(* IEC 61131-3 sources: IEC61131-3_ST_SCL_Mutation_Generator/Tests/mutatedCode_fibonacci_number_m, 23 files *)

(* ---- M1349.st ---- *)
FUNCTION_BLOCK "FB_Fibonacci_Calculator"
{ S7_Optimized_Access := 'FALSE' }
VERSION : 1.0

VAR_INPUT
    N : DInt := 5;
END_VAR

VAR_OUTPUT
    O : DInt := 1;
END_VAR

VAR
    F1 : DInt := 1;    // Fib(k-2) at the end of the calculation
    F2 : DInt := 1;    // Fib(k-1) at the end of the calculation
    CNT : DInt := 2;   // Index of the last computed term
END_VAR

BEGIN

    // Start values: Fib(1) = Fib(2) = 1
    #F1 := 1;
    #F2 := 1;
    #O := 1;

    IF #N >= 2 THEN (* MUTATED: REL_OP_REPLACE *)
        // Edge case: N <= 2 returns 1
        #CNT := #N;
    ELSE
        #CNT := 2;
        WHILE #CNT < #N DO
            #CNT := #CNT + 1;

            // Saturation arithmetic: result would exceed INT range
            IF (#F1 + #F2) > 32767 THEN
                #O := 32767;
                EXIT;
            END_IF;

            #O := #F1 + #F2;

            // Shift the window only if another term is still needed,
            // so that at the end O = F1 + F2
            IF #CNT < #N THEN
                #F1 := #F2;
                #F2 := #O;
            END_IF;
        END_WHILE;
    END_IF;

    // Final saturation guard
    IF (#O > 32767) OR (#O < 0) THEN
        #O := 32767;
    END_IF;

    //#ASSERT O >= 0 AND O <= 32767
    //#ASSERT F1 <= 32767 AND F2 <= 32767
    //#ASSERT CNT <= N

END_FUNCTION_BLOCK

(* ---- M1350.st ---- *)
FUNCTION_BLOCK "FB_Fibonacci_Calculator"
{ S7_Optimized_Access := 'FALSE' }
VERSION : 1.0

VAR_INPUT
    N : DInt := 5;
END_VAR

VAR_OUTPUT
    O : DInt := 1;
END_VAR

VAR
    F1 : DInt := 1;    // Fib(k-2) at the end of the calculation
    F2 : DInt := 1;    // Fib(k-1) at the end of the calculation
    CNT : DInt := 2;   // Index of the last computed term
END_VAR

BEGIN

    // Start values: Fib(1) = Fib(2) = 1
    #F1 := 1;
    #F2 := 1;
    #O := 1;

    IF #N <= 2 THEN
        // Edge case: N <= 2 returns 1
        #CNT := #N;
    ELSE
        #CNT := 2;
        WHILE #CNT > #N DO (* MUTATED: REL_OP_REPLACE *)
            #CNT := #CNT + 1;

            // Saturation arithmetic: result would exceed INT range
            IF (#F1 + #F2) > 32767 THEN
                #O := 32767;
                EXIT;
            END_IF;

            #O := #F1 + #F2;

            // Shift the window only if another term is still needed,
            // so that at the end O = F1 + F2
            IF #CNT < #N THEN
                #F1 := #F2;
                #F2 := #O;
            END_IF;
        END_WHILE;
    END_IF;

    // Final saturation guard
    IF (#O > 32767) OR (#O < 0) THEN
        #O := 32767;
    END_IF;

    //#ASSERT O >= 0 AND O <= 32767
    //#ASSERT F1 <= 32767 AND F2 <= 32767
    //#ASSERT CNT <= N

END_FUNCTION_BLOCK

(* ---- M1351.st ---- *)
FUNCTION_BLOCK "FB_Fibonacci_Calculator"
{ S7_Optimized_Access := 'FALSE' }
VERSION : 1.0

VAR_INPUT
    N : DInt := 5;
END_VAR

VAR_OUTPUT
    O : DInt := 1;
END_VAR

VAR
    F1 : DInt := 1;    // Fib(k-2) at the end of the calculation
    F2 : DInt := 1;    // Fib(k-1) at the end of the calculation
    CNT : DInt := 2;   // Index of the last computed term
END_VAR

BEGIN

    // Start values: Fib(1) = Fib(2) = 1
    #F1 := 1;
    #F2 := 1;
    #O := 1;

    IF #N <= 2 THEN
        // Edge case: N <= 2 returns 1
        #CNT := #N;
    ELSE
        #CNT := 2;
        WHILE #CNT < #N DO
            #CNT := #CNT + 1;

            // Saturation arithmetic: result would exceed INT range
            IF (#F1 + #F2) < 32767 THEN (* MUTATED: REL_OP_REPLACE *)
                #O := 32767;
                EXIT;
            END_IF;

            #O := #F1 + #F2;

            // Shift the window only if another term is still needed,
            // so that at the end O = F1 + F2
            IF #CNT < #N THEN
                #F1 := #F2;
                #F2 := #O;
            END_IF;
        END_WHILE;
    END_IF;

    // Final saturation guard
    IF (#O > 32767) OR (#O < 0) THEN
        #O := 32767;
    END_IF;

    //#ASSERT O >= 0 AND O <= 32767
    //#ASSERT F1 <= 32767 AND F2 <= 32767
    //#ASSERT CNT <= N

END_FUNCTION_BLOCK

(* ---- M1352.st ---- *)
FUNCTION_BLOCK "FB_Fibonacci_Calculator"
{ S7_Optimized_Access := 'FALSE' }
VERSION : 1.0

VAR_INPUT
    N : DInt := 5;
END_VAR

VAR_OUTPUT
    O : DInt := 1;
END_VAR

VAR
    F1 : DInt := 1;    // Fib(k-2) at the end of the calculation
    F2 : DInt := 1;    // Fib(k-1) at the end of the calculation
    CNT : DInt := 2;   // Index of the last computed term
END_VAR

BEGIN

    // Start values: Fib(1) = Fib(2) = 1
    #F1 := 1;
    #F2 := 1;
    #O := 1;

    IF #N <= 2 THEN
        // Edge case: N <= 2 returns 1
        #CNT := #N;
    ELSE
        #CNT := 2;
        WHILE #CNT < #N DO
            #CNT := #CNT + 1;

            // Saturation arithmetic: result would exceed INT range
            IF (#F1 + #F2) > 32767 THEN
                #O := 32767;
                EXIT;
            END_IF;

            #O := #F1 + #F2;

            // Shift the window only if another term is still needed,
            // so that at the end O = F1 + F2
            IF #CNT > #N THEN (* MUTATED: REL_OP_REPLACE *)
                #F1 := #F2;
                #F2 := #O;
            END_IF;
        END_WHILE;
    END_IF;

    // Final saturation guard
    IF (#O > 32767) OR (#O < 0) THEN
        #O := 32767;
    END_IF;

    //#ASSERT O >= 0 AND O <= 32767
    //#ASSERT F1 <= 32767 AND F2 <= 32767
    //#ASSERT CNT <= N

END_FUNCTION_BLOCK

(* ---- M1353.st ---- *)
FUNCTION_BLOCK "FB_Fibonacci_Calculator"
{ S7_Optimized_Access := 'FALSE' }
VERSION : 1.0

VAR_INPUT
    N : DInt := 5;
END_VAR

VAR_OUTPUT
    O : DInt := 1;
END_VAR

VAR
    F1 : DInt := 1;    // Fib(k-2) at the end of the calculation
    F2 : DInt := 1;    // Fib(k-1) at the end of the calculation
    CNT : DInt := 2;   // Index of the last computed term
END_VAR

BEGIN

    // Start values: Fib(1) = Fib(2) = 1
    #F1 := 1;
    #F2 := 1;
    #O := 1;

    IF #N <= 2 THEN
        // Edge case: N <= 2 returns 1
        #CNT := #N;
    ELSE
        #CNT := 2;
        WHILE #CNT < #N DO
            #CNT := #CNT + 1;

            // Saturation arithmetic: result would exceed INT range
            IF (#F1 + #F2) > 32767 THEN
                #O := 32767;
                EXIT;
            END_IF;

            #O := #F1 + #F2;

            // Shift the window only if another term is still needed,
            // so that at the end O = F1 + F2
            IF #CNT < #N THEN
                #F1 := #F2;
                #F2 := #O;
            END_IF;
        END_WHILE;
    END_IF;

    // Final saturation guard
    IF (#O < 32767) OR (#O < 0) THEN (* MUTATED: REL_OP_REPLACE *)
        #O := 32767;
    END_IF;

    //#ASSERT O >= 0 AND O <= 32767
    //#ASSERT F1 <= 32767 AND F2 <= 32767
    //#ASSERT CNT <= N

END_FUNCTION_BLOCK

(* ---- M1354.st ---- *)
FUNCTION_BLOCK "FB_Fibonacci_Calculator"
{ S7_Optimized_Access := 'FALSE' }
VERSION : 1.0

VAR_INPUT
    N : DInt := 5;
END_VAR

VAR_OUTPUT
    O : DInt := 1;
END_VAR

VAR
    F1 : DInt := 1;    // Fib(k-2) at the end of the calculation
    F2 : DInt := 1;    // Fib(k-1) at the end of the calculation
    CNT : DInt := 2;   // Index of the last computed term
END_VAR

BEGIN

    // Start values: Fib(1) = Fib(2) = 1
    #F1 := 1;
    #F2 := 1;
    #O := 1;

    IF #N <= 2 THEN
        // Edge case: N <= 2 returns 1
        #CNT := #N;
    ELSE
        #CNT := 2;
        WHILE #CNT < #N DO
            #CNT := #CNT + 1;

            // Saturation arithmetic: result would exceed INT range
            IF (#F1 + #F2) > 32767 THEN
                #O := 32767;
                EXIT;
            END_IF;

            #O := #F1 + #F2;

            // Shift the window only if another term is still needed,
            // so that at the end O = F1 + F2
            IF #CNT < #N THEN
                #F1 := #F2;
                #F2 := #O;
            END_IF;
        END_WHILE;
    END_IF;

    // Final saturation guard
    IF (#O > 32767) OR (#O > 0) THEN (* MUTATED: REL_OP_REPLACE *)
        #O := 32767;
    END_IF;

    //#ASSERT O >= 0 AND O <= 32767
    //#ASSERT F1 <= 32767 AND F2 <= 32767
    //#ASSERT CNT <= N

END_FUNCTION_BLOCK

(* ---- M1355.st ---- *)
FUNCTION_BLOCK "FB_Fibonacci_Calculator"
{ S7_Optimized_Access := 'FALSE' }
VERSION : 1.0

VAR_INPUT
    N : DInt := 5;
END_VAR

VAR_OUTPUT
    O : DInt := 1;
END_VAR

VAR
    F1 : DInt := 1;    // Fib(k-2) at the end of the calculation
    F2 : DInt := 1;    // Fib(k-1) at the end of the calculation
    CNT : DInt := 2;   // Index of the last computed term
END_VAR

BEGIN

    // Start values: Fib(1) = Fib(2) = 1
    #F1 := 1;
    #F2 := 1;
    #O := 1;

    IF #N <= 2 THEN
        // Edge case: N <= 2 returns 1
        #CNT := #N;
    ELSE
        #CNT := 2;
        WHILE #CNT < #N DO
            #CNT := #CNT + 1;

            // Saturation arithmetic: result would exceed INT range
            IF (#F1 + #F2) > 32767 THEN
                #O := 32767;
                EXIT;
            END_IF;

            #O := #F1 + #F2;

            // Shift the window only if another term is still needed,
            // so that at the end O = F1 + F2
            IF #CNT < #N THEN
                #F1 := #F2;
                #F2 := #O;
            END_IF;
        END_WHILE;
    END_IF;

    // Final saturation guard
    IF (#O > 32767) AND (#O < 0) THEN (* MUTATED: LOGICAL_OP_REPLACE *)
        #O := 32767;
    END_IF;

    //#ASSERT O >= 0 AND O <= 32767
    //#ASSERT F1 <= 32767 AND F2 <= 32767
    //#ASSERT CNT <= N

END_FUNCTION_BLOCK

(* ---- M1356.st ---- *)
FUNCTION_BLOCK "FB_Fibonacci_Calculator"
{ S7_Optimized_Access := 'FALSE' }
VERSION : 1.0

VAR_INPUT
    N : DInt := 5;
END_VAR

VAR_OUTPUT
    O : DInt := 1;
END_VAR

VAR
    F1 : DInt := 1;    // Fib(k-2) at the end of the calculation
    F2 : DInt := 1;    // Fib(k-1) at the end of the calculation
    CNT : DInt := 2;   // Index of the last computed term
END_VAR

BEGIN

    // Start values: Fib(1) = Fib(2) = 1
    #F1 := 1;
    #F2 := 1;
    #O := 1;

    IF #N <= 2 THEN
        // Edge case: N <= 2 returns 1
        #CNT := #N;
    ELSE
        #CNT := 2;
        WHILE #CNT < #N DO
            #CNT := #CNT - 1; (* MUTATED: ARITH_OP_REPLACE *)

            // Saturation arithmetic: result would exceed INT range
            IF (#F1 + #F2) > 32767 THEN
                #O := 32767;
                EXIT;
            END_IF;

            #O := #F1 + #F2;

            // Shift the window only if another term is still needed,
            // so that at the end O = F1 + F2
            IF #CNT < #N THEN
                #F1 := #F2;
                #F2 := #O;
            END_IF;
        END_WHILE;
    END_IF;

    // Final saturation guard
    IF (#O > 32767) OR (#O < 0) THEN
        #O := 32767;
    END_IF;

    //#ASSERT O >= 0 AND O <= 32767
    //#ASSERT F1 <= 32767 AND F2 <= 32767
    //#ASSERT CNT <= N

END_FUNCTION_BLOCK

(* ---- M1357.st ---- *)
FUNCTION_BLOCK "FB_Fibonacci_Calculator"
{ S7_Optimized_Access := 'FALSE' }
VERSION : 1.0

VAR_INPUT
    N : DInt := 5;
END_VAR

VAR_OUTPUT
    O : DInt := 1;
END_VAR

VAR
    F1 : DInt := 1;    // Fib(k-2) at the end of the calculation
    F2 : DInt := 1;    // Fib(k-1) at the end of the calculation
    CNT : DInt := 2;   // Index of the last computed term
END_VAR

BEGIN

    // Start values: Fib(1) = Fib(2) = 1
    #F1 := 2; (* MUTATED: CONST_VALUE_REPLACE *)
    #F2 := 1;
    #O := 1;

    IF #N <= 2 THEN
        // Edge case: N <= 2 returns 1
        #CNT := #N;
    ELSE
        #CNT := 2;
        WHILE #CNT < #N DO
            #CNT := #CNT + 1;

            // Saturation arithmetic: result would exceed INT range
            IF (#F1 + #F2) > 32767 THEN
                #O := 32767;
                EXIT;
            END_IF;

            #O := #F1 + #F2;

            // Shift the window only if another term is still needed,
            // so that at the end O = F1 + F2
            IF #CNT < #N THEN
                #F1 := #F2;
                #F2 := #O;
            END_IF;
        END_WHILE;
    END_IF;

    // Final saturation guard
    IF (#O > 32767) OR (#O < 0) THEN
        #O := 32767;
    END_IF;

    //#ASSERT O >= 0 AND O <= 32767
    //#ASSERT F1 <= 32767 AND F2 <= 32767
    //#ASSERT CNT <= N

END_FUNCTION_BLOCK

(* ---- M1358.st ---- *)
FUNCTION_BLOCK "FB_Fibonacci_Calculator"
{ S7_Optimized_Access := 'FALSE' }
VERSION : 1.0

VAR_INPUT
    N : DInt := 5;
END_VAR

VAR_OUTPUT
    O : DInt := 1;
END_VAR

VAR
    F1 : DInt := 1;    // Fib(k-2) at the end of the calculation
    F2 : DInt := 1;    // Fib(k-1) at the end of the calculation
    CNT : DInt := 2;   // Index of the last computed term
END_VAR

BEGIN

    // Start values: Fib(1) = Fib(2) = 1
    #F1 := 1;
    #F2 := 2; (* MUTATED: CONST_VALUE_REPLACE *)
    #O := 1;

    IF #N <= 2 THEN
        // Edge case: N <= 2 returns 1
        #CNT := #N;
    ELSE
        #CNT := 2;
        WHILE #CNT < #N DO
            #CNT := #CNT + 1;

            // Saturation arithmetic: result would exceed INT range
            IF (#F1 + #F2) > 32767 THEN
                #O := 32767;
                EXIT;
            END_IF;

            #O := #F1 + #F2;

            // Shift the window only if another term is still needed,
            // so that at the end O = F1 + F2
            IF #CNT < #N THEN
                #F1 := #F2;
                #F2 := #O;
            END_IF;
        END_WHILE;
    END_IF;

    // Final saturation guard
    IF (#O > 32767) OR (#O < 0) THEN
        #O := 32767;
    END_IF;

    //#ASSERT O >= 0 AND O <= 32767
    //#ASSERT F1 <= 32767 AND F2 <= 32767
    //#ASSERT CNT <= N

END_FUNCTION_BLOCK

(* ---- M1359.st ---- *)
FUNCTION_BLOCK "FB_Fibonacci_Calculator"
{ S7_Optimized_Access := 'FALSE' }
VERSION : 1.0

VAR_INPUT
    N : DInt := 5;
END_VAR

VAR_OUTPUT
    O : DInt := 1;
END_VAR

VAR
    F1 : DInt := 1;    // Fib(k-2) at the end of the calculation
    F2 : DInt := 1;    // Fib(k-1) at the end of the calculation
    CNT : DInt := 2;   // Index of the last computed term
END_VAR

BEGIN

    // Start values: Fib(1) = Fib(2) = 1
    #F1 := 1;
    #F2 := 1;
    #O := 2; (* MUTATED: CONST_VALUE_REPLACE *)

    IF #N <= 2 THEN
        // Edge case: N <= 2 returns 1
        #CNT := #N;
    ELSE
        #CNT := 2;
        WHILE #CNT < #N DO
            #CNT := #CNT + 1;

            // Saturation arithmetic: result would exceed INT range
            IF (#F1 + #F2) > 32767 THEN
                #O := 32767;
                EXIT;
            END_IF;

            #O := #F1 + #F2;

            // Shift the window only if another term is still needed,
            // so that at the end O = F1 + F2
            IF #CNT < #N THEN
                #F1 := #F2;
                #F2 := #O;
            END_IF;
        END_WHILE;
    END_IF;

    // Final saturation guard
    IF (#O > 32767) OR (#O < 0) THEN
        #O := 32767;
    END_IF;

    //#ASSERT O >= 0 AND O <= 32767
    //#ASSERT F1 <= 32767 AND F2 <= 32767
    //#ASSERT CNT <= N

END_FUNCTION_BLOCK

(* ---- M1360.st ---- *)
FUNCTION_BLOCK "FB_Fibonacci_Calculator"
{ S7_Optimized_Access := 'FALSE' }
VERSION : 1.0

VAR_INPUT
    N : DInt := 5;
END_VAR

VAR_OUTPUT
    O : DInt := 1;
END_VAR

VAR
    F1 : DInt := 1;    // Fib(k-2) at the end of the calculation
    F2 : DInt := 1;    // Fib(k-1) at the end of the calculation
    CNT : DInt := 2;   // Index of the last computed term
END_VAR

BEGIN

    // Start values: Fib(1) = Fib(2) = 1
    #F1 := 1;
    #F2 := 1;
    #O := 1;

    IF #N <= 3 THEN (* MUTATED: CONST_VALUE_REPLACE *)
        // Edge case: N <= 2 returns 1
        #CNT := #N;
    ELSE
        #CNT := 2;
        WHILE #CNT < #N DO
            #CNT := #CNT + 1;

            // Saturation arithmetic: result would exceed INT range
            IF (#F1 + #F2) > 32767 THEN
                #O := 32767;
                EXIT;
            END_IF;

            #O := #F1 + #F2;

            // Shift the window only if another term is still needed,
            // so that at the end O = F1 + F2
            IF #CNT < #N THEN
                #F1 := #F2;
                #F2 := #O;
            END_IF;
        END_WHILE;
    END_IF;

    // Final saturation guard
    IF (#O > 32767) OR (#O < 0) THEN
        #O := 32767;
    END_IF;

    //#ASSERT O >= 0 AND O <= 32767
    //#ASSERT F1 <= 32767 AND F2 <= 32767
    //#ASSERT CNT <= N

END_FUNCTION_BLOCK

(* ---- M1361.st ---- *)
FUNCTION_BLOCK "FB_Fibonacci_Calculator"
{ S7_Optimized_Access := 'FALSE' }
VERSION : 1.0

VAR_INPUT
    N : DInt := 5;
END_VAR

VAR_OUTPUT
    O : DInt := 1;
END_VAR

VAR
    F1 : DInt := 1;    // Fib(k-2) at the end of the calculation
    F2 : DInt := 1;    // Fib(k-1) at the end of the calculation
    CNT : DInt := 2;   // Index of the last computed term
END_VAR

BEGIN

    // Start values: Fib(1) = Fib(2) = 1
    #F1 := 1;
    #F2 := 1;
    #O := 1;

    IF #N <= 2 THEN
        // Edge case: N <= 2 returns 1
        #CNT := #N;
    ELSE
        #CNT := 3; (* MUTATED: CONST_VALUE_REPLACE *)
        WHILE #CNT < #N DO
            #CNT := #CNT + 1;

            // Saturation arithmetic: result would exceed INT range
            IF (#F1 + #F2) > 32767 THEN
                #O := 32767;
                EXIT;
            END_IF;

            #O := #F1 + #F2;

            // Shift the window only if another term is still needed,
            // so that at the end O = F1 + F2
            IF #CNT < #N THEN
                #F1 := #F2;
                #F2 := #O;
            END_IF;
        END_WHILE;
    END_IF;

    // Final saturation guard
    IF (#O > 32767) OR (#O < 0) THEN
        #O := 32767;
    END_IF;

    //#ASSERT O >= 0 AND O <= 32767
    //#ASSERT F1 <= 32767 AND F2 <= 32767
    //#ASSERT CNT <= N

END_FUNCTION_BLOCK

(* ---- M1362.st ---- *)
FUNCTION_BLOCK "FB_Fibonacci_Calculator"
{ S7_Optimized_Access := 'FALSE' }
VERSION : 1.0

VAR_INPUT
    N : DInt := 5;
END_VAR

VAR_OUTPUT
    O : DInt := 1;
END_VAR

VAR
    F1 : DInt := 1;    // Fib(k-2) at the end of the calculation
    F2 : DInt := 1;    // Fib(k-1) at the end of the calculation
    CNT : DInt := 2;   // Index of the last computed term
END_VAR

BEGIN

    // Start values: Fib(1) = Fib(2) = 1
    #F1 := 1;
    #F2 := 1;
    #O := 1;

    IF #N <= 2 THEN
        // Edge case: N <= 2 returns 1
        #CNT := #N;
    ELSE
        #CNT := 2;
        WHILE #CNT < #N DO
            #CNT := #CNT + 2; (* MUTATED: CONST_VALUE_REPLACE *)

            // Saturation arithmetic: result would exceed INT range
            IF (#F1 + #F2) > 32767 THEN
                #O := 32767;
                EXIT;
            END_IF;

            #O := #F1 + #F2;

            // Shift the window only if another term is still needed,
            // so that at the end O = F1 + F2
            IF #CNT < #N THEN
                #F1 := #F2;
                #F2 := #O;
            END_IF;
        END_WHILE;
    END_IF;

    // Final saturation guard
    IF (#O > 32767) OR (#O < 0) THEN
        #O := 32767;
    END_IF;

    //#ASSERT O >= 0 AND O <= 32767
    //#ASSERT F1 <= 32767 AND F2 <= 32767
    //#ASSERT CNT <= N

END_FUNCTION_BLOCK

(* ---- M1363.st ---- *)
FUNCTION_BLOCK "FB_Fibonacci_Calculator"
{ S7_Optimized_Access := 'FALSE' }
VERSION : 1.0

VAR_INPUT
    N : DInt := 5;
END_VAR

VAR_OUTPUT
    O : DInt := 1;
END_VAR

VAR
    F1 : DInt := 1;    // Fib(k-2) at the end of the calculation
    F2 : DInt := 1;    // Fib(k-1) at the end of the calculation
    CNT : DInt := 2;   // Index of the last computed term
END_VAR

BEGIN

    // Start values: Fib(1) = Fib(2) = 1
    #F1 := 1;
    #F2 := 1;
    #O := 1;

    IF #N <= 2 THEN
        // Edge case: N <= 2 returns 1
        #CNT := #N;
    ELSE
        #CNT := 2;
        WHILE #CNT < #N DO
            #CNT := #CNT + 1;

            // Saturation arithmetic: result would exceed INT range
            IF (#F1 + #F2) > 32768 THEN (* MUTATED: CONST_VALUE_REPLACE *)
                #O := 32767;
                EXIT;
            END_IF;

            #O := #F1 + #F2;

            // Shift the window only if another term is still needed,
            // so that at the end O = F1 + F2
            IF #CNT < #N THEN
                #F1 := #F2;
                #F2 := #O;
            END_IF;
        END_WHILE;
    END_IF;

    // Final saturation guard
    IF (#O > 32767) OR (#O < 0) THEN
        #O := 32767;
    END_IF;

    //#ASSERT O >= 0 AND O <= 32767
    //#ASSERT F1 <= 32767 AND F2 <= 32767
    //#ASSERT CNT <= N

END_FUNCTION_BLOCK

(* ---- M1364.st ---- *)
FUNCTION_BLOCK "FB_Fibonacci_Calculator"
{ S7_Optimized_Access := 'FALSE' }
VERSION : 1.0

VAR_INPUT
    N : DInt := 5;
END_VAR

VAR_OUTPUT
    O : DInt := 1;
END_VAR

VAR
    F1 : DInt := 1;    // Fib(k-2) at the end of the calculation
    F2 : DInt := 1;    // Fib(k-1) at the end of the calculation
    CNT : DInt := 2;   // Index of the last computed term
END_VAR

BEGIN

    // Start values: Fib(1) = Fib(2) = 1
    #F1 := 1;
    #F2 := 1;
    #O := 1;

    IF #N <= 2 THEN
        // Edge case: N <= 2 returns 1
        #CNT := #N;
    ELSE
        #CNT := 2;
        WHILE #CNT < #N DO
            #CNT := #CNT + 1;

            // Saturation arithmetic: result would exceed INT range
            IF (#F1 + #F2) > 32767 THEN
                #O := 32768; (* MUTATED: CONST_VALUE_REPLACE *)
                EXIT;
            END_IF;

            #O := #F1 + #F2;

            // Shift the window only if another term is still needed,
            // so that at the end O = F1 + F2
            IF #CNT < #N THEN
                #F1 := #F2;
                #F2 := #O;
            END_IF;
        END_WHILE;
    END_IF;

    // Final saturation guard
    IF (#O > 32767) OR (#O < 0) THEN
        #O := 32767;
    END_IF;

    //#ASSERT O >= 0 AND O <= 32767
    //#ASSERT F1 <= 32767 AND F2 <= 32767
    //#ASSERT CNT <= N

END_FUNCTION_BLOCK

(* ---- M1365.st ---- *)
FUNCTION_BLOCK "FB_Fibonacci_Calculator"
{ S7_Optimized_Access := 'FALSE' }
VERSION : 1.0

VAR_INPUT
    N : DInt := 5;
END_VAR

VAR_OUTPUT
    O : DInt := 1;
END_VAR

VAR
    F1 : DInt := 1;    // Fib(k-2) at the end of the calculation
    F2 : DInt := 1;    // Fib(k-1) at the end of the calculation
    CNT : DInt := 2;   // Index of the last computed term
END_VAR

BEGIN

    // Start values: Fib(1) = Fib(2) = 1
    #F1 := 1;
    #F2 := 1;
    #O := 1;

    IF #N <= 2 THEN
        // Edge case: N <= 2 returns 1
        #CNT := #N;
    ELSE
        #CNT := 2;
        WHILE #CNT < #N DO
            #CNT := #CNT + 1;

            // Saturation arithmetic: result would exceed INT range
            IF (#F1 + #F2) > 32767 THEN
                #O := 32767;
                EXIT;
            END_IF;

            #O := #F1 + #F2;

            // Shift the window only if another term is still needed,
            // so that at the end O = F1 + F2
            IF #CNT < #N THEN
                #F1 := #F2;
                #F2 := #O;
            END_IF;
        END_WHILE;
    END_IF;

    // Final saturation guard
    IF (#O > 32768) OR (#O < 0) THEN (* MUTATED: CONST_VALUE_REPLACE *)
        #O := 32767;
    END_IF;

    //#ASSERT O >= 0 AND O <= 32767
    //#ASSERT F1 <= 32767 AND F2 <= 32767
    //#ASSERT CNT <= N

END_FUNCTION_BLOCK

(* ---- M1366.st ---- *)
FUNCTION_BLOCK "FB_Fibonacci_Calculator"
{ S7_Optimized_Access := 'FALSE' }
VERSION : 1.0

VAR_INPUT
    N : DInt := 5;
END_VAR

VAR_OUTPUT
    O : DInt := 1;
END_VAR

VAR
    F1 : DInt := 1;    // Fib(k-2) at the end of the calculation
    F2 : DInt := 1;    // Fib(k-1) at the end of the calculation
    CNT : DInt := 2;   // Index of the last computed term
END_VAR

BEGIN

    // Start values: Fib(1) = Fib(2) = 1
    #F1 := 1;
    #F2 := 1;
    #O := 1;

    IF #N <= 2 THEN
        // Edge case: N <= 2 returns 1
        #CNT := #N;
    ELSE
        #CNT := 2;
        WHILE #CNT < #N DO
            #CNT := #CNT + 1;

            // Saturation arithmetic: result would exceed INT range
            IF (#F1 + #F2) > 32767 THEN
                #O := 32767;
                EXIT;
            END_IF;

            #O := #F1 + #F2;

            // Shift the window only if another term is still needed,
            // so that at the end O = F1 + F2
            IF #CNT < #N THEN
                #F1 := #F2;
                #F2 := #O;
            END_IF;
        END_WHILE;
    END_IF;

    // Final saturation guard
    IF (#O > 32767) OR (#O < 1) THEN (* MUTATED: CONST_VALUE_REPLACE *)
        #O := 32767;
    END_IF;

    //#ASSERT O >= 0 AND O <= 32767
    //#ASSERT F1 <= 32767 AND F2 <= 32767
    //#ASSERT CNT <= N

END_FUNCTION_BLOCK

(* ---- M1367.st ---- *)
FUNCTION_BLOCK "FB_Fibonacci_Calculator"
{ S7_Optimized_Access := 'FALSE' }
VERSION : 1.0

VAR_INPUT
    N : DInt := 5;
END_VAR

VAR_OUTPUT
    O : DInt := 1;
END_VAR

VAR
    F1 : DInt := 1;    // Fib(k-2) at the end of the calculation
    F2 : DInt := 1;    // Fib(k-1) at the end of the calculation
    CNT : DInt := 2;   // Index of the last computed term
END_VAR

BEGIN

    // Start values: Fib(1) = Fib(2) = 1
    #F1 := 1;
    #F2 := 1;
    #O := 1;

    IF #N <= 2 THEN
        // Edge case: N <= 2 returns 1
        #CNT := #N;
    ELSE
        #CNT := 2;
        WHILE #CNT < #N DO
            #CNT := #CNT + 1;

            // Saturation arithmetic: result would exceed INT range
            IF (#F1 + #F2) > 32767 THEN
                #O := 32767;
                EXIT;
            END_IF;

            #O := #F1 + #F2;

            // Shift the window only if another term is still needed,
            // so that at the end O = F1 + F2
            IF #CNT < #N THEN
                #F1 := #F2;
                #F2 := #O;
            END_IF;
        END_WHILE;
    END_IF;

    // Final saturation guard
    IF (#O > 32767) OR (#O < 0) THEN
        #O := 32768; (* MUTATED: CONST_VALUE_REPLACE *)
    END_IF;

    //#ASSERT O >= 0 AND O <= 32767
    //#ASSERT F1 <= 32767 AND F2 <= 32767
    //#ASSERT CNT <= N

END_FUNCTION_BLOCK

(* ---- M1368.st ---- *)
FUNCTION_BLOCK "FB_Fibonacci_Calculator"
{ S7_Optimized_Access := 'FALSE' }
VERSION : 1.0

VAR_INPUT
    N : DInt := 5;
END_VAR

VAR_OUTPUT
    O : DInt := 1;
END_VAR

VAR
    F1 : DInt := 1;    // Fib(k-2) at the end of the calculation
    F2 : DInt := 1;    // Fib(k-1) at the end of the calculation
    CNT : DInt := 2;   // Index of the last computed term
END_VAR

BEGIN

    // Start values: Fib(1) = Fib(2) = 1
    #F1 := 1;
    #F2 := 1;
    #O := 1;

    IF NOT (#N <= 2) THEN (* MUTATED: COND_NEGATE *)
        // Edge case: N <= 2 returns 1
        #CNT := #N;
    ELSE
        #CNT := 2;
        WHILE #CNT < #N DO
            #CNT := #CNT + 1;

            // Saturation arithmetic: result would exceed INT range
            IF (#F1 + #F2) > 32767 THEN
                #O := 32767;
                EXIT;
            END_IF;

            #O := #F1 + #F2;

            // Shift the window only if another term is still needed,
            // so that at the end O = F1 + F2
            IF #CNT < #N THEN
                #F1 := #F2;
                #F2 := #O;
            END_IF;
        END_WHILE;
    END_IF;

    // Final saturation guard
    IF (#O > 32767) OR (#O < 0) THEN
        #O := 32767;
    END_IF;

    //#ASSERT O >= 0 AND O <= 32767
    //#ASSERT F1 <= 32767 AND F2 <= 32767
    //#ASSERT CNT <= N

END_FUNCTION_BLOCK

(* ---- M1369.st ---- *)
FUNCTION_BLOCK "FB_Fibonacci_Calculator"
{ S7_Optimized_Access := 'FALSE' }
VERSION : 1.0

VAR_INPUT
    N : DInt := 5;
END_VAR

VAR_OUTPUT
    O : DInt := 1;
END_VAR

VAR
    F1 : DInt := 1;    // Fib(k-2) at the end of the calculation
    F2 : DInt := 1;    // Fib(k-1) at the end of the calculation
    CNT : DInt := 2;   // Index of the last computed term
END_VAR

BEGIN

    // Start values: Fib(1) = Fib(2) = 1
    #F1 := 1;
    #F2 := 1;
    #O := 1;

    IF #N <= 2 THEN
        // Edge case: N <= 2 returns 1
        #CNT := #N;
    ELSE
        #CNT := 2;
        WHILE #CNT < #N DO
            #CNT := #CNT + 1;

            // Saturation arithmetic: result would exceed INT range
            IF NOT ((#F1 + #F2) > 32767) THEN (* MUTATED: COND_NEGATE *)
                #O := 32767;
                EXIT;
            END_IF;

            #O := #F1 + #F2;

            // Shift the window only if another term is still needed,
            // so that at the end O = F1 + F2
            IF #CNT < #N THEN
                #F1 := #F2;
                #F2 := #O;
            END_IF;
        END_WHILE;
    END_IF;

    // Final saturation guard
    IF (#O > 32767) OR (#O < 0) THEN
        #O := 32767;
    END_IF;

    //#ASSERT O >= 0 AND O <= 32767
    //#ASSERT F1 <= 32767 AND F2 <= 32767
    //#ASSERT CNT <= N

END_FUNCTION_BLOCK

(* ---- M1370.st ---- *)
FUNCTION_BLOCK "FB_Fibonacci_Calculator"
{ S7_Optimized_Access := 'FALSE' }
VERSION : 1.0

VAR_INPUT
    N : DInt := 5;
END_VAR

VAR_OUTPUT
    O : DInt := 1;
END_VAR

VAR
    F1 : DInt := 1;    // Fib(k-2) at the end of the calculation
    F2 : DInt := 1;    // Fib(k-1) at the end of the calculation
    CNT : DInt := 2;   // Index of the last computed term
END_VAR

BEGIN

    // Start values: Fib(1) = Fib(2) = 1
    #F1 := 1;
    #F2 := 1;
    #O := 1;

    IF #N <= 2 THEN
        // Edge case: N <= 2 returns 1
        #CNT := #N;
    ELSE
        #CNT := 2;
        WHILE #CNT < #N DO
            #CNT := #CNT + 1;

            // Saturation arithmetic: result would exceed INT range
            IF (#F1 + #F2) > 32767 THEN
                #O := 32767;
                EXIT;
            END_IF;

            #O := #F1 + #F2;

            // Shift the window only if another term is still needed,
            // so that at the end O = F1 + F2
            IF NOT (#CNT < #N) THEN (* MUTATED: COND_NEGATE *)
                #F1 := #F2;
                #F2 := #O;
            END_IF;
        END_WHILE;
    END_IF;

    // Final saturation guard
    IF (#O > 32767) OR (#O < 0) THEN
        #O := 32767;
    END_IF;

    //#ASSERT O >= 0 AND O <= 32767
    //#ASSERT F1 <= 32767 AND F2 <= 32767
    //#ASSERT CNT <= N

END_FUNCTION_BLOCK

(* ---- M1371.st ---- *)
FUNCTION_BLOCK "FB_Fibonacci_Calculator"
{ S7_Optimized_Access := 'FALSE' }
VERSION : 1.0

VAR_INPUT
    N : DInt := 5;
END_VAR

VAR_OUTPUT
    O : DInt := 1;
END_VAR

VAR
    F1 : DInt := 1;    // Fib(k-2) at the end of the calculation
    F2 : DInt := 1;    // Fib(k-1) at the end of the calculation
    CNT : DInt := 2;   // Index of the last computed term
END_VAR

BEGIN

    // Start values: Fib(1) = Fib(2) = 1
    #F1 := 1;
    #F2 := 1;
    #O := 1;

    IF #N <= 2 THEN
        // Edge case: N <= 2 returns 1
        #CNT := #N;
    ELSE
        #CNT := 2;
        WHILE #CNT < #N DO
            #CNT := #CNT + 1;

            // Saturation arithmetic: result would exceed INT range
            IF (#F1 + #F2) > 32767 THEN
                #O := 32767;
                EXIT;
            END_IF;

            #O := #F1 + #F2;

            // Shift the window only if another term is still needed,
            // so that at the end O = F1 + F2
            IF #CNT < #N THEN
                #F1 := #F2;
                #F2 := #O;
            END_IF;
        END_WHILE;
    END_IF;

    // Final saturation guard
    IF NOT ((#O > 32767) OR (#O < 0)) THEN (* MUTATED: COND_NEGATE *)
        #O := 32767;
    END_IF;

    //#ASSERT O >= 0 AND O <= 32767
    //#ASSERT F1 <= 32767 AND F2 <= 32767
    //#ASSERT CNT <= N

END_FUNCTION_BLOCK
